(* IEC 61131-3 sources: ironplc/compiler/sources/resources/libs/Tc2_System/1.0.0, 1 file *)

(* ---- Tc2_System.st ---- *)
(* Tc2_System compatibility library -- global constants.

   This file reproduces the *interface* (the constant name PI and its value)
   of Beckhoff's TwinCAT Tc2_System library for interoperability. IronPLC is an
   independent open-source project and is not affiliated with, endorsed by, or
   sponsored by Beckhoff Automation GmbH. See
   specs/steering/compatibility-library-authoring.md. *)
VAR_GLOBAL CONSTANT
    PI : LREAL := 3.1415926535897932384626433832795;
END_VAR
